Fanuc KAREL source: kc00008.KL

-- PROVISIONAL review KL for V770-1; original PC SHA256 8fd84556a8a24b9ed4e3b41106443df11bc7407ddb581a1056505731256aa37d
-- Incomplete behavior may be omitted. Consult companion uncertainty JSON. Do not deploy.
PROGRAM KC00008
%NOLOCKGROUP
BEGIN
  -- UNRESOLVED_PC offsets 5-33; opcodes 27,22,1C,22,22,31
  -- UNRESOLVED_PC offsets 38-42; opcodes 7F
END KC00008
